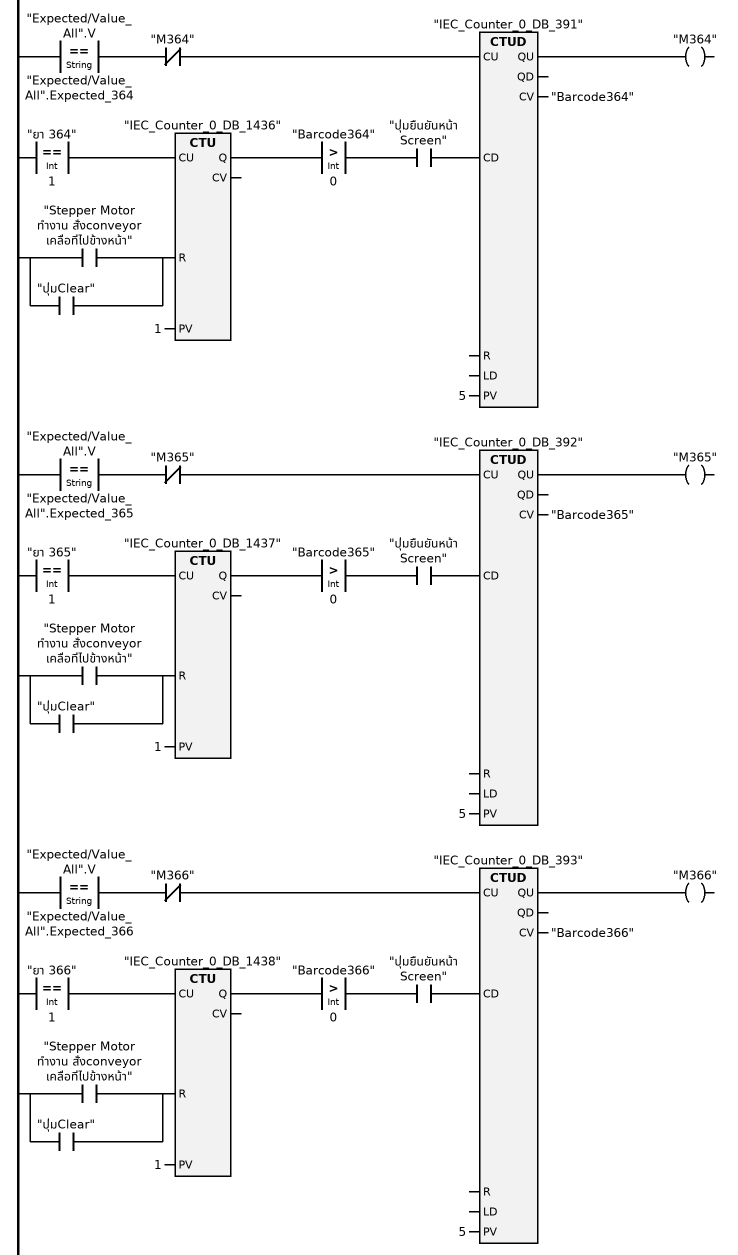
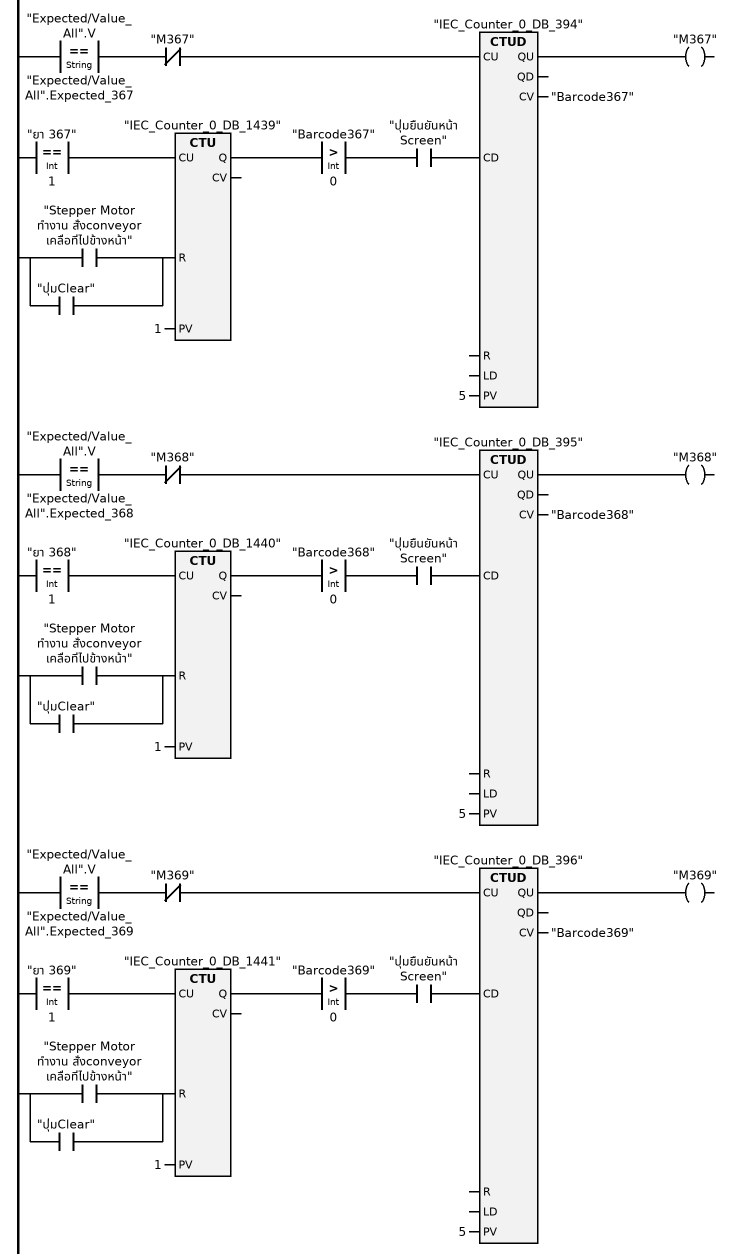
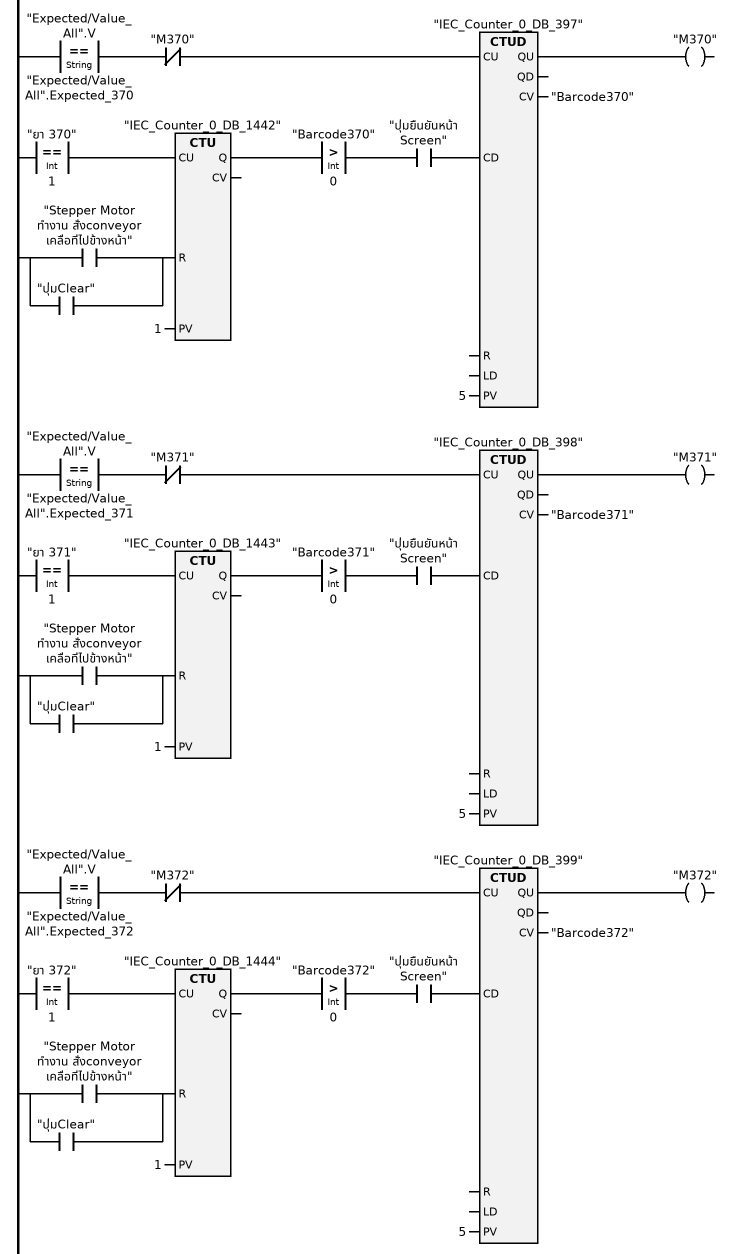
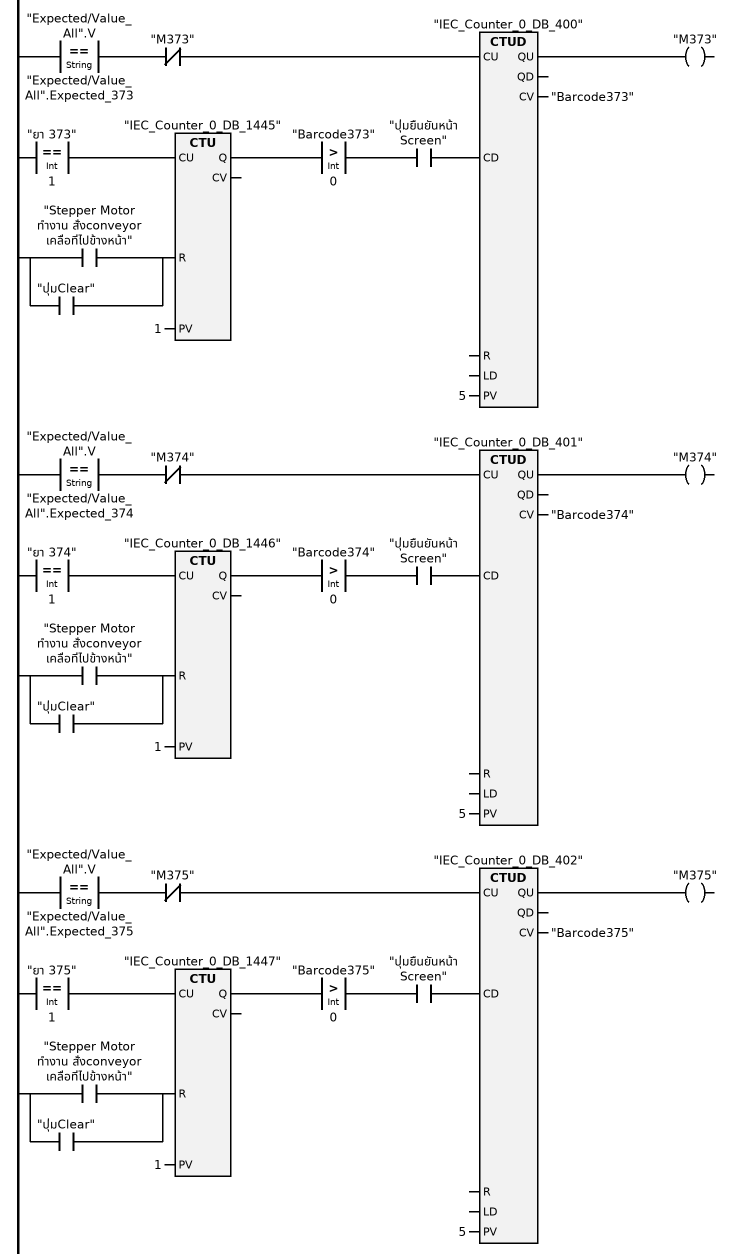
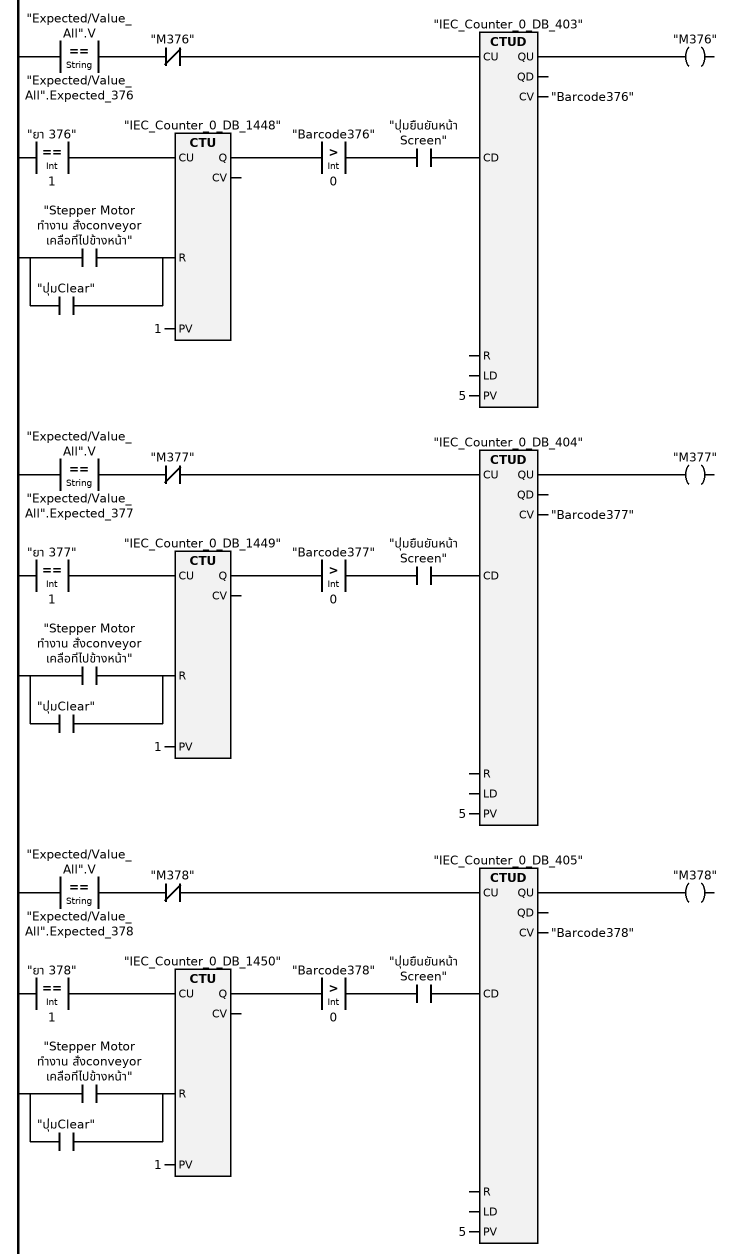
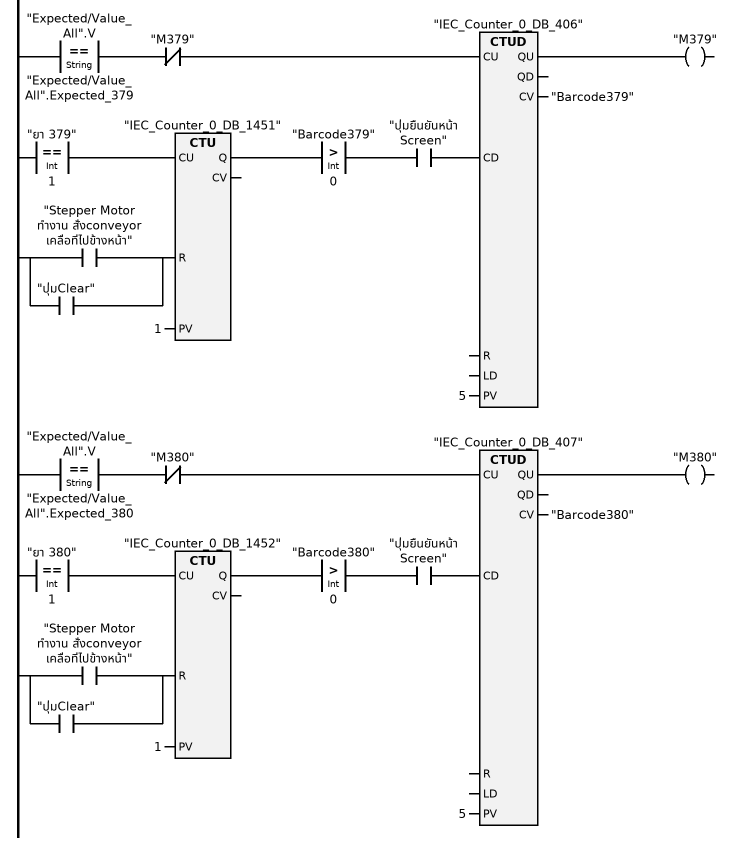
   "IEC_Counter_0_DB_1433".CTU(CU := "ยา 361" = 1,
                           R := "Stepper Motor ทำงาน สั่งconveyor เคลื่อที่ไปข้างหน้า" OR "ปุ่มClear",
                           PV := 1);
   "IEC_Counter_0_DB_388".CTUD(CU := ("Expected/Value_All".V = "Expected/Value_All".Expected_361) AND NOT "M361",
                           CD := "IEC_Counter_0_DB_1433".Q AND ("Barcode361" > 0) AND "ปุ่มยืนยันหน้า Screen",
                           PV := 5,
                           CV => "Barcode361");
   "M361" := "IEC_Counter_0_DB_388".QU;
   "IEC_Counter_0_DB_1434".CTU(CU := "ยา 362" = 1,
                           R := "Stepper Motor ทำงาน สั่งconveyor เคลื่อที่ไปข้างหน้า" OR "ปุ่มClear",
                           PV := 1);
   "IEC_Counter_0_DB_389".CTUD(CU := ("Expected/Value_All".V = "Expected/Value_All".Expected_362) AND NOT "M362",
                           CD := "IEC_Counter_0_DB_1434".Q AND ("Barcode362" > 0) AND "ปุ่มยืนยันหน้า Screen",
                           PV := 5,
                           CV => "Barcode362");
   "M362" := "IEC_Counter_0_DB_389".QU;
   "IEC_Counter_0_DB_1435".CTU(CU := "ยา 363" = 1,
                           R := "Stepper Motor ทำงาน สั่งconveyor เคลื่อที่ไปข้างหน้า" OR "ปุ่มClear",
                           PV := 1);
   "IEC_Counter_0_DB_390".CTUD(CU := ("Expected/Value_All".V = "Expected/Value_All".Expected_363) AND NOT "M363",
                           CD := "IEC_Counter_0_DB_1435".Q AND ("Barcode363" > 0) AND "ปุ่มยืนยันหน้า Screen",
                           PV := 5,
                           CV => "Barcode363");
   "M363" := "IEC_Counter_0_DB_390".QU;
   "IEC_Counter_0_DB_1436".CTU(CU := "ยา 364" = 1,
                           R := "Stepper Motor ทำงาน สั่งconveyor เคลื่อที่ไปข้างหน้า" OR "ปุ่มClear",
                           PV := 1);
   "IEC_Counter_0_DB_391".CTUD(CU := ("Expected/Value_All".V = "Expected/Value_All".Expected_364) AND NOT "M364",
                           CD := "IEC_Counter_0_DB_1436".Q AND ("Barcode364" > 0) AND "ปุ่มยืนยันหน้า Screen",
                           PV := 5,
                           CV => "Barcode364");
   "M364" := "IEC_Counter_0_DB_391".QU;
   "IEC_Counter_0_DB_1437".CTU(CU := "ยา 365" = 1,
                           R := "Stepper Motor ทำงาน สั่งconveyor เคลื่อที่ไปข้างหน้า" OR "ปุ่มClear",
                           PV := 1);
   "IEC_Counter_0_DB_392".CTUD(CU := ("Expected/Value_All".V = "Expected/Value_All".Expected_365) AND NOT "M365",
                           CD := "IEC_Counter_0_DB_1437".Q AND ("Barcode365" > 0) AND "ปุ่มยืนยันหน้า Screen",
                           PV := 5,
                           CV => "Barcode365");
   "M365" := "IEC_Counter_0_DB_392".QU;
   "IEC_Counter_0_DB_1438".CTU(CU := "ยา 366" = 1,
                           R := "Stepper Motor ทำงาน สั่งconveyor เคลื่อที่ไปข้างหน้า" OR "ปุ่มClear",
                           PV := 1);
   "IEC_Counter_0_DB_393".CTUD(CU := ("Expected/Value_All".V = "Expected/Value_All".Expected_366) AND NOT "M366",
                           CD := "IEC_Counter_0_DB_1438".Q AND ("Barcode366" > 0) AND "ปุ่มยืนยันหน้า Screen",
                           PV := 5,
                           CV => "Barcode366");
   "M366" := "IEC_Counter_0_DB_393".QU;
   "IEC_Counter_0_DB_1439".CTU(CU := "ยา 367" = 1,
                           R := "Stepper Motor ทำงาน สั่งconveyor เคลื่อที่ไปข้างหน้า" OR "ปุ่มClear",
                           PV := 1);
   "IEC_Counter_0_DB_394".CTUD(CU := ("Expected/Value_All".V = "Expected/Value_All".Expected_367) AND NOT "M367",
                           CD := "IEC_Counter_0_DB_1439".Q AND ("Barcode367" > 0) AND "ปุ่มยืนยันหน้า Screen",
                           PV := 5,
                           CV => "Barcode367");
   "M367" := "IEC_Counter_0_DB_394".QU;
   "IEC_Counter_0_DB_1440".CTU(CU := "ยา 368" = 1,
                           R := "Stepper Motor ทำงาน สั่งconveyor เคลื่อที่ไปข้างหน้า" OR "ปุ่มClear",
                           PV := 1);
   "IEC_Counter_0_DB_395".CTUD(CU := ("Expected/Value_All".V = "Expected/Value_All".Expected_368) AND NOT "M368",
                           CD := "IEC_Counter_0_DB_1440".Q AND ("Barcode368" > 0) AND "ปุ่มยืนยันหน้า Screen",
                           PV := 5,
                           CV => "Barcode368");
   "M368" := "IEC_Counter_0_DB_395".QU;
   "IEC_Counter_0_DB_1441".CTU(CU := "ยา 369" = 1,
                           R := "Stepper Motor ทำงาน สั่งconveyor เคลื่อที่ไปข้างหน้า" OR "ปุ่มClear",
                           PV := 1);
   "IEC_Counter_0_DB_396".CTUD(CU := ("Expected/Value_All".V = "Expected/Value_All".Expected_369) AND NOT "M369",
                           CD := "IEC_Counter_0_DB_1441".Q AND ("Barcode369" > 0) AND "ปุ่มยืนยันหน้า Screen",
                           PV := 5,
                           CV => "Barcode369");
   "M369" := "IEC_Counter_0_DB_396".QU;
   "IEC_Counter_0_DB_1442".CTU(CU := "ยา 370" = 1,
                           R := "Stepper Motor ทำงาน สั่งconveyor เคลื่อที่ไปข้างหน้า" OR "ปุ่มClear",
                           PV := 1);
   "IEC_Counter_0_DB_397".CTUD(CU := ("Expected/Value_All".V = "Expected/Value_All".Expected_370) AND NOT "M370",
                           CD := "IEC_Counter_0_DB_1442".Q AND ("Barcode370" > 0) AND "ปุ่มยืนยันหน้า Screen",
                           PV := 5,
                           CV => "Barcode370");
   "M370" := "IEC_Counter_0_DB_397".QU;
   "IEC_Counter_0_DB_1443".CTU(CU := "ยา 371" = 1,
                           R := "Stepper Motor ทำงาน สั่งconveyor เคลื่อที่ไปข้างหน้า" OR "ปุ่มClear",
                           PV := 1);
   "IEC_Counter_0_DB_398".CTUD(CU := ("Expected/Value_All".V = "Expected/Value_All".Expected_371) AND NOT "M371",
                           CD := "IEC_Counter_0_DB_1443".Q AND ("Barcode371" > 0) AND "ปุ่มยืนยันหน้า Screen",
                           PV := 5,
                           CV => "Barcode371");
   "M371" := "IEC_Counter_0_DB_398".QU;
   "IEC_Counter_0_DB_1444".CTU(CU := "ยา 372" = 1,
                           R := "Stepper Motor ทำงาน สั่งconveyor เคลื่อที่ไปข้างหน้า" OR "ปุ่มClear",
                           PV := 1);
   "IEC_Counter_0_DB_399".CTUD(CU := ("Expected/Value_All".V = "Expected/Value_All".Expected_372) AND NOT "M372",
                           CD := "IEC_Counter_0_DB_1444".Q AND ("Barcode372" > 0) AND "ปุ่มยืนยันหน้า Screen",
                           PV := 5,
                           CV => "Barcode372");
   "M372" := "IEC_Counter_0_DB_399".QU;
   "IEC_Counter_0_DB_1445".CTU(CU := "ยา 373" = 1,
                           R := "Stepper Motor ทำงาน สั่งconveyor เคลื่อที่ไปข้างหน้า" OR "ปุ่มClear",
                           PV := 1);
   "IEC_Counter_0_DB_400".CTUD(CU := ("Expected/Value_All".V = "Expected/Value_All".Expected_373) AND NOT "M373",
                           CD := "IEC_Counter_0_DB_1445".Q AND ("Barcode373" > 0) AND "ปุ่มยืนยันหน้า Screen",
                           PV := 5,
                           CV => "Barcode373");
   "M373" := "IEC_Counter_0_DB_400".QU;
   "IEC_Counter_0_DB_1446".CTU(CU := "ยา 374" = 1,
                           R := "Stepper Motor ทำงาน สั่งconveyor เคลื่อที่ไปข้างหน้า" OR "ปุ่มClear",
                           PV := 1);
   "IEC_Counter_0_DB_401".CTUD(CU := ("Expected/Value_All".V = "Expected/Value_All".Expected_374) AND NOT "M374",
                           CD := "IEC_Counter_0_DB_1446".Q AND ("Barcode374" > 0) AND "ปุ่มยืนยันหน้า Screen",
                           PV := 5,
                           CV => "Barcode374");
   "M374" := "IEC_Counter_0_DB_401".QU;
   "IEC_Counter_0_DB_1447".CTU(CU := "ยา 375" = 1,
                           R := "Stepper Motor ทำงาน สั่งconveyor เคลื่อที่ไปข้างหน้า" OR "ปุ่มClear",
                           PV := 1);
   "IEC_Counter_0_DB_402".CTUD(CU := ("Expected/Value_All".V = "Expected/Value_All".Expected_375) AND NOT "M375",
                           CD := "IEC_Counter_0_DB_1447".Q AND ("Barcode375" > 0) AND "ปุ่มยืนยันหน้า Screen",
                           PV := 5,
                           CV => "Barcode375");
   "M375" := "IEC_Counter_0_DB_402".QU;
   "IEC_Counter_0_DB_1448".CTU(CU := "ยา 376" = 1,
                           R := "Stepper Motor ทำงาน สั่งconveyor เคลื่อที่ไปข้างหน้า" OR "ปุ่มClear",
                           PV := 1);
   "IEC_Counter_0_DB_403".CTUD(CU := ("Expected/Value_All".V = "Expected/Value_All".Expected_376) AND NOT "M376",
                           CD := "IEC_Counter_0_DB_1448".Q AND ("Barcode376" > 0) AND "ปุ่มยืนยันหน้า Screen",
                           PV := 5,
                           CV => "Barcode376");
   "M376" := "IEC_Counter_0_DB_403".QU;
   "IEC_Counter_0_DB_1449".CTU(CU := "ยา 377" = 1,
                           R := "Stepper Motor ทำงาน สั่งconveyor เคลื่อที่ไปข้างหน้า" OR "ปุ่มClear",
                           PV := 1);
   "IEC_Counter_0_DB_404".CTUD(CU := ("Expected/Value_All".V = "Expected/Value_All".Expected_377) AND NOT "M377",
                           CD := "IEC_Counter_0_DB_1449".Q AND ("Barcode377" > 0) AND "ปุ่มยืนยันหน้า Screen",
                           PV := 5,
                           CV => "Barcode377");
   "M377" := "IEC_Counter_0_DB_404".QU;
   "IEC_Counter_0_DB_1450".CTU(CU := "ยา 378" = 1,
                           R := "Stepper Motor ทำงาน สั่งconveyor เคลื่อที่ไปข้างหน้า" OR "ปุ่มClear",
                           PV := 1);
   "IEC_Counter_0_DB_405".CTUD(CU := ("Expected/Value_All".V = "Expected/Value_All".Expected_378) AND NOT "M378",
                           CD := "IEC_Counter_0_DB_1450".Q AND ("Barcode378" > 0) AND "ปุ่มยืนยันหน้า Screen",
                           PV := 5,
                           CV => "Barcode378");
   "M378" := "IEC_Counter_0_DB_405".QU;
   "IEC_Counter_0_DB_1451".CTU(CU := "ยา 379" = 1,
                           R := "Stepper Motor ทำงาน สั่งconveyor เคลื่อที่ไปข้างหน้า" OR "ปุ่มClear",
                           PV := 1);
   "IEC_Counter_0_DB_406".CTUD(CU := ("Expected/Value_All".V = "Expected/Value_All".Expected_379) AND NOT "M379",
                           CD := "IEC_Counter_0_DB_1451".Q AND ("Barcode379" > 0) AND "ปุ่มยืนยันหน้า Screen",
                           PV := 5,
                           CV => "Barcode379");
   "M379" := "IEC_Counter_0_DB_406".QU;
   "IEC_Counter_0_DB_1452".CTU(CU := "ยา 380" = 1,
                           R := "Stepper Motor ทำงาน สั่งconveyor เคลื่อที่ไปข้างหน้า" OR "ปุ่มClear",
                           PV := 1);
   "IEC_Counter_0_DB_407".CTUD(CU := ("Expected/Value_All".V = "Expected/Value_All".Expected_380) AND NOT "M380",
                           CD := "IEC_Counter_0_DB_1452".Q AND ("Barcode380" > 0) AND "ปุ่มยืนยันหน้า Screen",
                           PV := 5,
                           CV => "Barcode380");
   "M380" := "IEC_Counter_0_DB_407".QU;
END_REGION

REGION Network 20
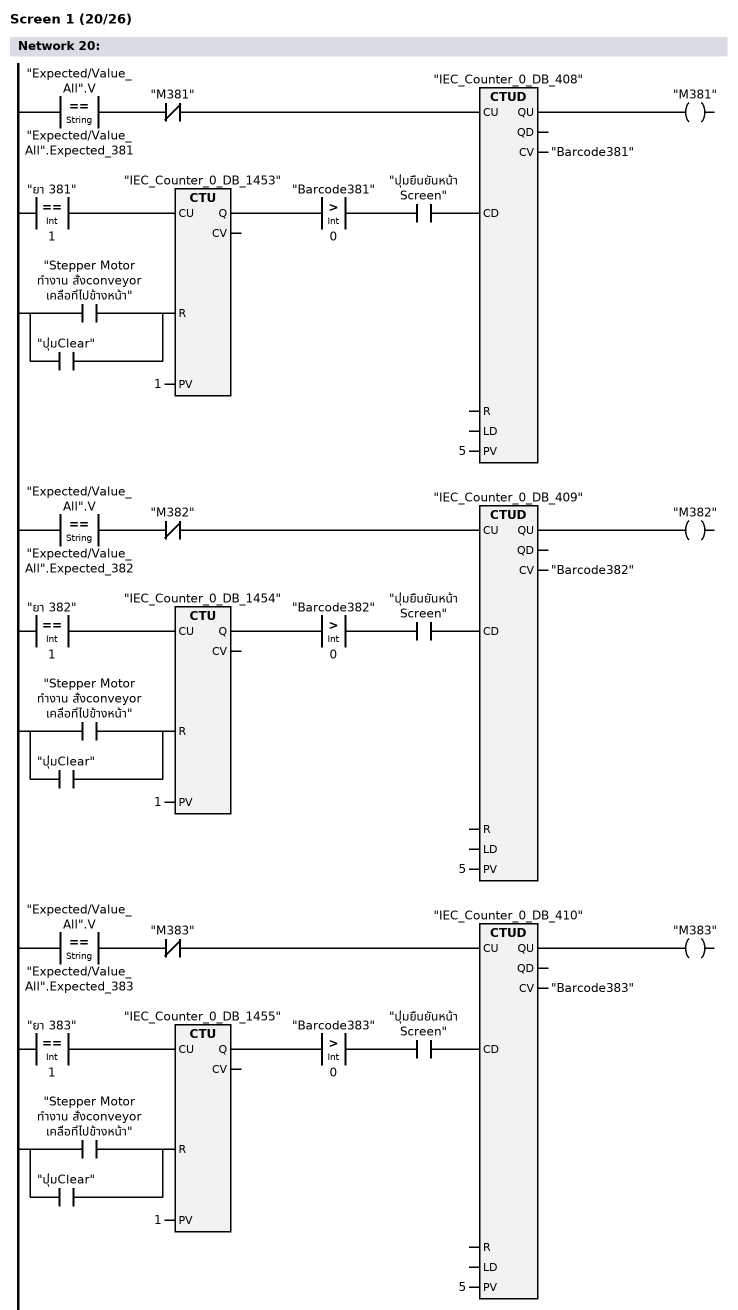
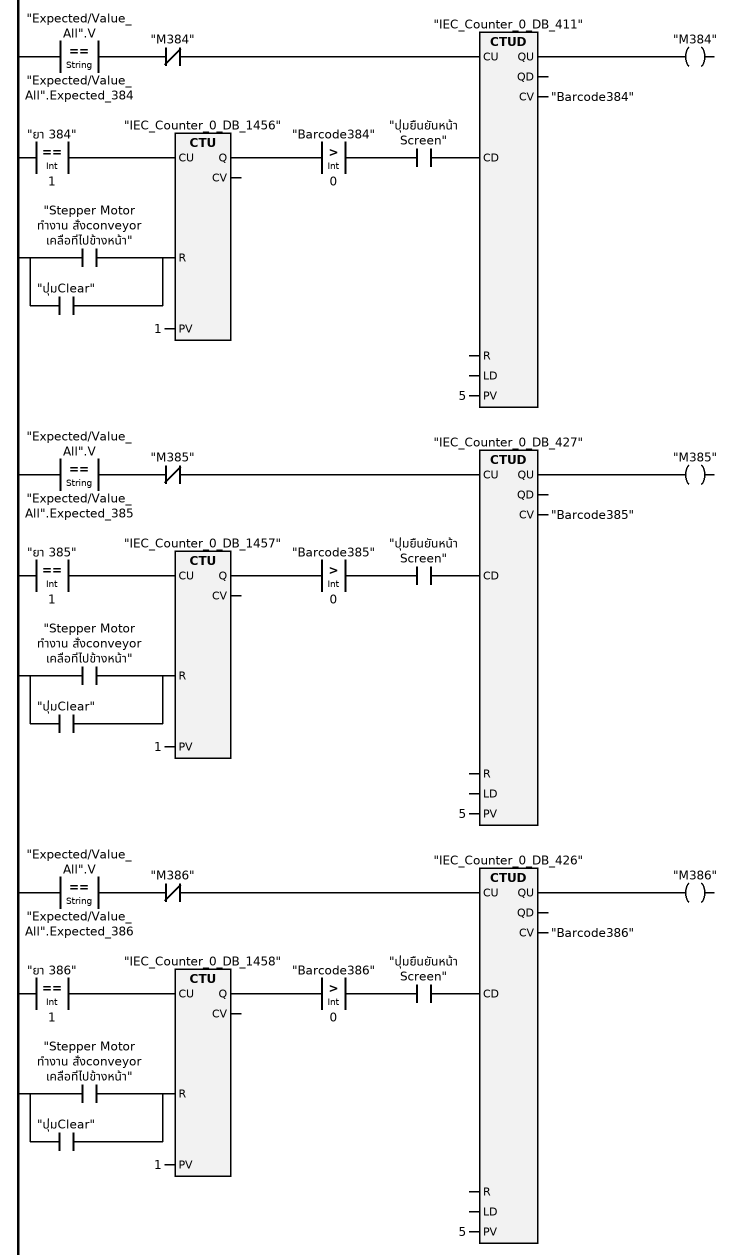
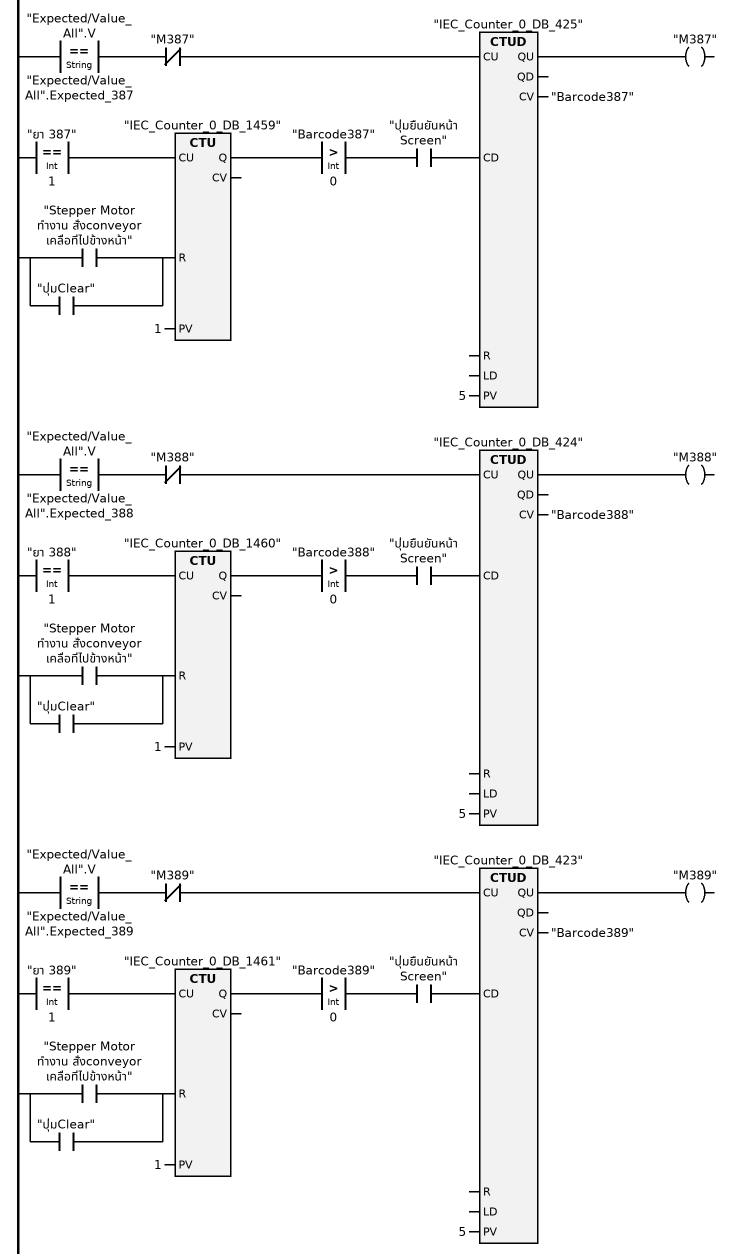
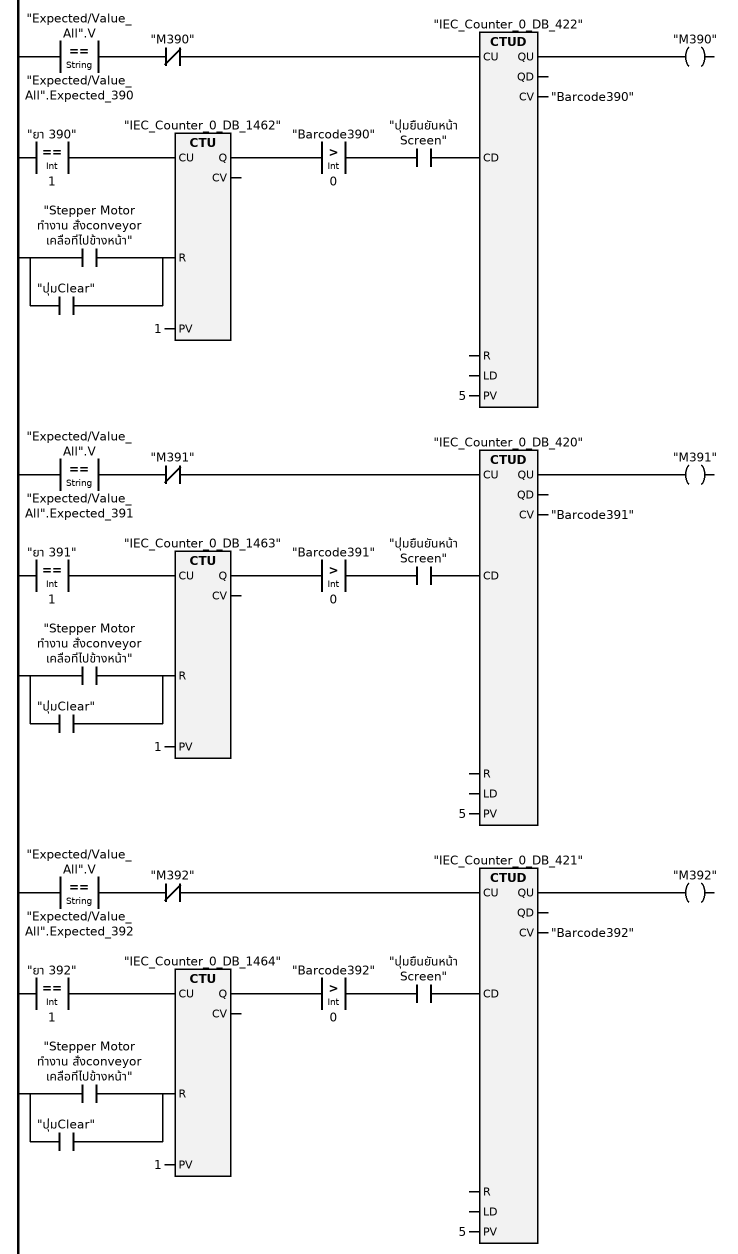
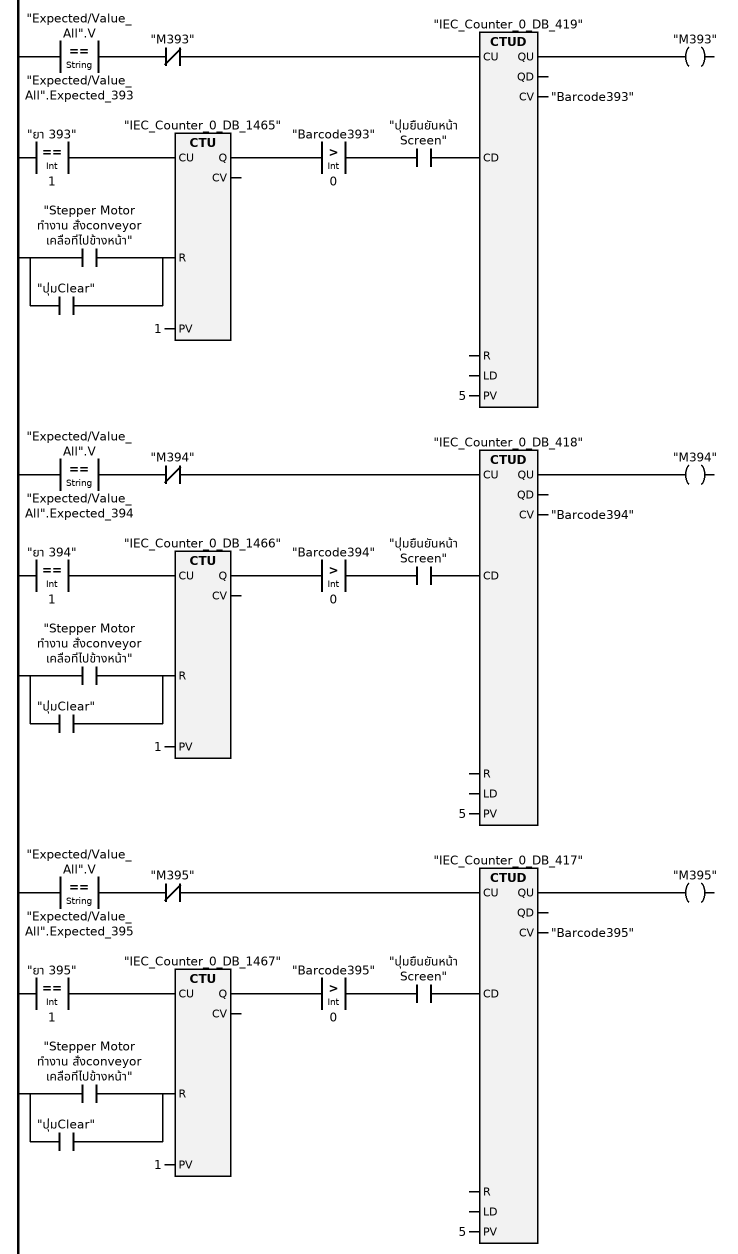
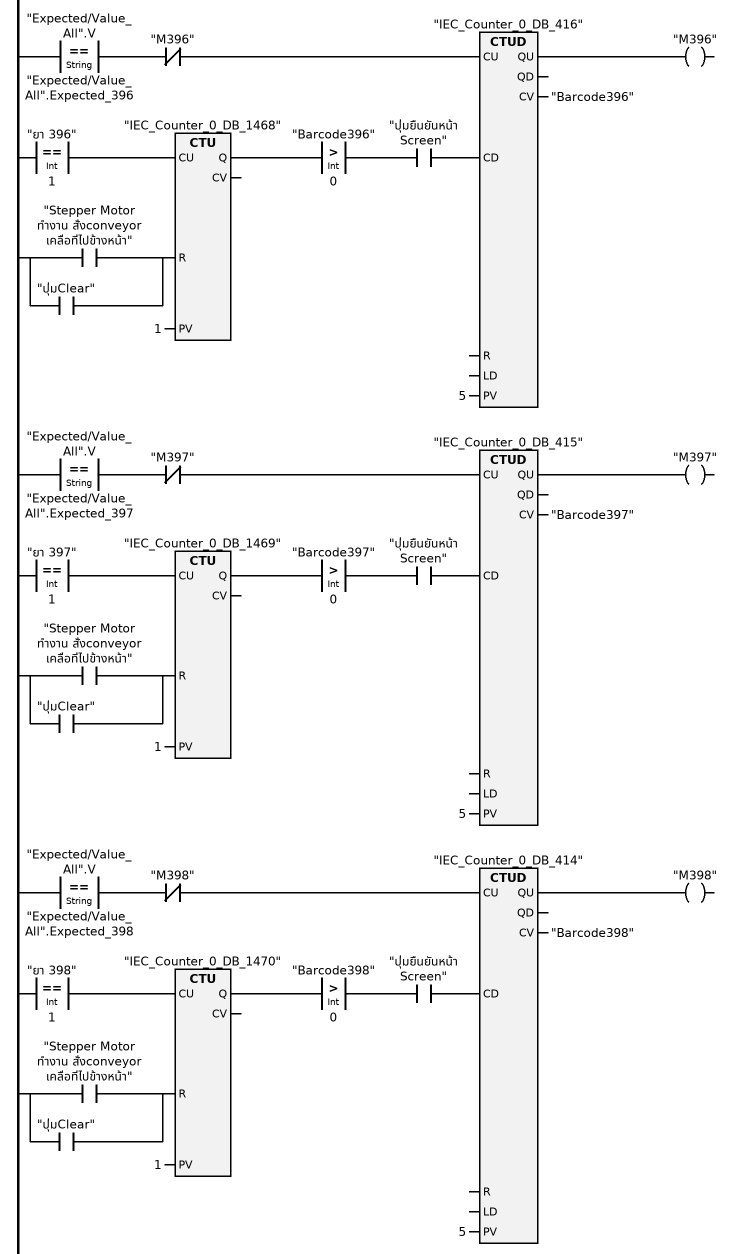
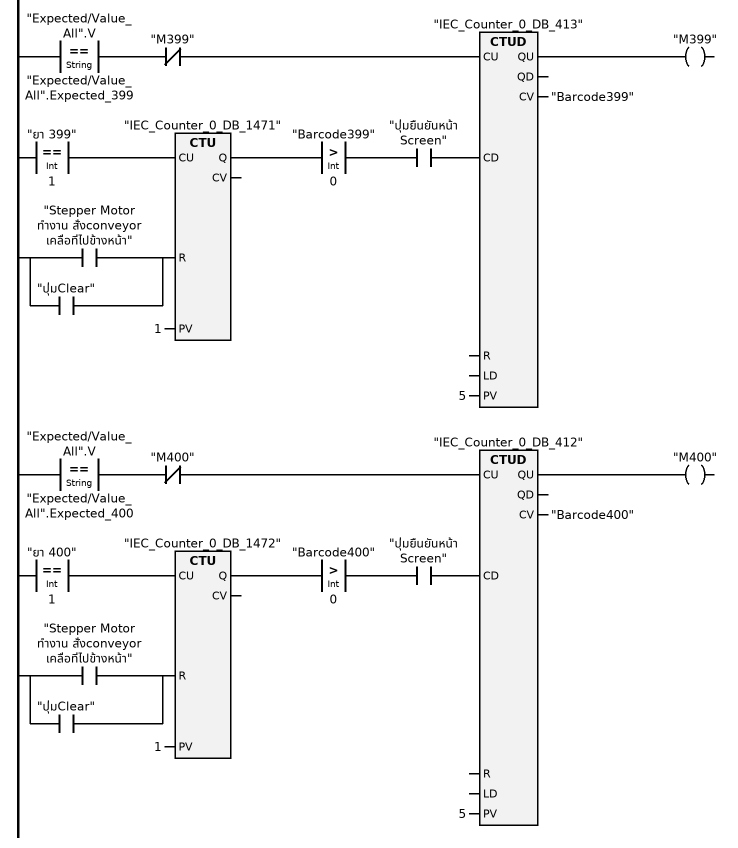
   "IEC_Counter_0_DB_1453".CTU(CU := "ยา 381" = 1,
                           R := "Stepper Motor ทำงาน สั่งconveyor เคลื่อที่ไปข้างหน้า" OR "ปุ่มClear",
                           PV := 1);
   "IEC_Counter_0_DB_408".CTUD(CU := ("Expected/Value_All".V = "Expected/Value_All".Expected_381) AND NOT "M381",
                           CD := "IEC_Counter_0_DB_1453".Q AND ("Barcode381" > 0) AND "ปุ่มยืนยันหน้า Screen",
                           PV := 5,
                           CV => "Barcode381");
   "M381" := "IEC_Counter_0_DB_408".QU;
   "IEC_Counter_0_DB_1454".CTU(CU := "ยา 382" = 1,
                           R := "Stepper Motor ทำงาน สั่งconveyor เคลื่อที่ไปข้างหน้า" OR "ปุ่มClear",
                           PV := 1);
   "IEC_Counter_0_DB_409".CTUD(CU := ("Expected/Value_All".V = "Expected/Value_All".Expected_382) AND NOT "M382",
                           CD := "IEC_Counter_0_DB_1454".Q AND ("Barcode382" > 0) AND "ปุ่มยืนยันหน้า Screen",
                           PV := 5,
                           CV => "Barcode382");
   "M382" := "IEC_Counter_0_DB_409".QU;
   "IEC_Counter_0_DB_1455".CTU(CU := "ยา 383" = 1,
                           R := "Stepper Motor ทำงาน สั่งconveyor เคลื่อที่ไปข้างหน้า" OR "ปุ่มClear",
                           PV := 1);
   "IEC_Counter_0_DB_410".CTUD(CU := ("Expected/Value_All".V = "Expected/Value_All".Expected_383) AND NOT "M383",
                           CD := "IEC_Counter_0_DB_1455".Q AND ("Barcode383" > 0) AND "ปุ่มยืนยันหน้า Screen",
                           PV := 5,
                           CV => "Barcode383");
   "M383" := "IEC_Counter_0_DB_410".QU;
   "IEC_Counter_0_DB_1456".CTU(CU := "ยา 384" = 1,
                           R := "Stepper Motor ทำงาน สั่งconveyor เคลื่อที่ไปข้างหน้า" OR "ปุ่มClear",
                           PV := 1);
   "IEC_Counter_0_DB_411".CTUD(CU := ("Expected/Value_All".V = "Expected/Value_All".Expected_384) AND NOT "M384",
                           CD := "IEC_Counter_0_DB_1456".Q AND ("Barcode384" > 0) AND "ปุ่มยืนยันหน้า Screen",
                           PV := 5,
                           CV => "Barcode384");
   "M384" := "IEC_Counter_0_DB_411".QU;
   "IEC_Counter_0_DB_1457".CTU(CU := "ยา 385" = 1,
                           R := "Stepper Motor ทำงาน สั่งconveyor เคลื่อที่ไปข้างหน้า" OR "ปุ่มClear",
                           PV := 1);
   "IEC_Counter_0_DB_427".CTUD(CU := ("Expected/Value_All".V = "Expected/Value_All".Expected_385) AND NOT "M385",
                           CD := "IEC_Counter_0_DB_1457".Q AND ("Barcode385" > 0) AND "ปุ่มยืนยันหน้า Screen",
                           PV := 5,
                           CV => "Barcode385");
   "M385" := "IEC_Counter_0_DB_427".QU;
   "IEC_Counter_0_DB_1458".CTU(CU := "ยา 386" = 1,
                           R := "Stepper Motor ทำงาน สั่งconveyor เคลื่อที่ไปข้างหน้า" OR "ปุ่มClear",
                           PV := 1);
   "IEC_Counter_0_DB_426".CTUD(CU := ("Expected/Value_All".V = "Expected/Value_All".Expected_386) AND NOT "M386",
                           CD := "IEC_Counter_0_DB_1458".Q AND ("Barcode386" > 0) AND "ปุ่มยืนยันหน้า Screen",
                           PV := 5,
                           CV => "Barcode386");
   "M386" := "IEC_Counter_0_DB_426".QU;
   "IEC_Counter_0_DB_1459".CTU(CU := "ยา 387" = 1,
                           R := "Stepper Motor ทำงาน สั่งconveyor เคลื่อที่ไปข้างหน้า" OR "ปุ่มClear",
                           PV := 1);
   "IEC_Counter_0_DB_425".CTUD(CU := ("Expected/Value_All".V = "Expected/Value_All".Expected_387) AND NOT "M387",
                           CD := "IEC_Counter_0_DB_1459".Q AND ("Barcode387" > 0) AND "ปุ่มยืนยันหน้า Screen",
                           PV := 5,
                           CV => "Barcode387");
   "M387" := "IEC_Counter_0_DB_425".QU;
   "IEC_Counter_0_DB_1460".CTU(CU := "ยา 388" = 1,
                           R := "Stepper Motor ทำงาน สั่งconveyor เคลื่อที่ไปข้างหน้า" OR "ปุ่มClear",
                           PV := 1);
   "IEC_Counter_0_DB_424".CTUD(CU := ("Expected/Value_All".V = "Expected/Value_All".Expected_388) AND NOT "M388",
                           CD := "IEC_Counter_0_DB_1460".Q AND ("Barcode388" > 0) AND "ปุ่มยืนยันหน้า Screen",
                           PV := 5,
                           CV => "Barcode388");
   "M388" := "IEC_Counter_0_DB_424".QU;
   "IEC_Counter_0_DB_1461".CTU(CU := "ยา 389" = 1,
                           R := "Stepper Motor ทำงาน สั่งconveyor เคลื่อที่ไปข้างหน้า" OR "ปุ่มClear",
                           PV := 1);
   "IEC_Counter_0_DB_423".CTUD(CU := ("Expected/Value_All".V = "Expected/Value_All".Expected_389) AND NOT "M389",
                           CD := "IEC_Counter_0_DB_1461".Q AND ("Barcode389" > 0) AND "ปุ่มยืนยันหน้า Screen",
                           PV := 5,
                           CV => "Barcode389");
   "M389" := "IEC_Counter_0_DB_423".QU;
   "IEC_Counter_0_DB_1462".CTU(CU := "ยา 390" = 1,
                           R := "Stepper Motor ทำงาน สั่งconveyor เคลื่อที่ไปข้างหน้า" OR "ปุ่มClear",
                           PV := 1);
   "IEC_Counter_0_DB_422".CTUD(CU := ("Expected/Value_All".V = "Expected/Value_All".Expected_390) AND NOT "M390",
                           CD := "IEC_Counter_0_DB_1462".Q AND ("Barcode390" > 0) AND "ปุ่มยืนยันหน้า Screen",
                           PV := 5,
                           CV => "Barcode390");
   "M390" := "IEC_Counter_0_DB_422".QU;
   "IEC_Counter_0_DB_1463".CTU(CU := "ยา 391" = 1,
                           R := "Stepper Motor ทำงาน สั่งconveyor เคลื่อที่ไปข้างหน้า" OR "ปุ่มClear",
                           PV := 1);
   "IEC_Counter_0_DB_420".CTUD(CU := ("Expected/Value_All".V = "Expected/Value_All".Expected_391) AND NOT "M391",
                           CD := "IEC_Counter_0_DB_1463".Q AND ("Barcode391" > 0) AND "ปุ่มยืนยันหน้า Screen",
                           PV := 5,
                           CV => "Barcode391");
   "M391" := "IEC_Counter_0_DB_420".QU;
   "IEC_Counter_0_DB_1464".CTU(CU := "ยา 392" = 1,
                           R := "Stepper Motor ทำงาน สั่งconveyor เคลื่อที่ไปข้างหน้า" OR "ปุ่มClear",
                           PV := 1);
   "IEC_Counter_0_DB_421".CTUD(CU := ("Expected/Value_All".V = "Expected/Value_All".Expected_392) AND NOT "M392",
                           CD := "IEC_Counter_0_DB_1464".Q AND ("Barcode392" > 0) AND "ปุ่มยืนยันหน้า Screen",
                           PV := 5,
                           CV => "Barcode392");
   "M392" := "IEC_Counter_0_DB_421".QU;
   "IEC_Counter_0_DB_1465".CTU(CU := "ยา 393" = 1,
                           R := "Stepper Motor ทำงาน สั่งconveyor เคลื่อที่ไปข้างหน้า" OR "ปุ่มClear",
                           PV := 1);
   "IEC_Counter_0_DB_419".CTUD(CU := ("Expected/Value_All".V = "Expected/Value_All".Expected_393) AND NOT "M393",
                           CD := "IEC_Counter_0_DB_1465".Q AND ("Barcode393" > 0) AND "ปุ่มยืนยันหน้า Screen",
                           PV := 5,
                           CV => "Barcode393");
   "M393" := "IEC_Counter_0_DB_419".QU;
   "IEC_Counter_0_DB_1466".CTU(CU := "ยา 394" = 1,
                           R := "Stepper Motor ทำงาน สั่งconveyor เคลื่อที่ไปข้างหน้า" OR "ปุ่มClear",
                           PV := 1);
   "IEC_Counter_0_DB_418".CTUD(CU := ("Expected/Value_All".V = "Expected/Value_All".Expected_394) AND NOT "M394",
                           CD := "IEC_Counter_0_DB_1466".Q AND ("Barcode394" > 0) AND "ปุ่มยืนยันหน้า Screen",
                           PV := 5,
                           CV => "Barcode394");
   "M394" := "IEC_Counter_0_DB_418".QU;
   "IEC_Counter_0_DB_1467".CTU(CU := "ยา 395" = 1,
                           R := "Stepper Motor ทำงาน สั่งconveyor เคลื่อที่ไปข้างหน้า" OR "ปุ่มClear",
                           PV := 1);
   "IEC_Counter_0_DB_417".CTUD(CU := ("Expected/Value_All".V = "Expected/Value_All".Expected_395) AND NOT "M395",
                           CD := "IEC_Counter_0_DB_1467".Q AND ("Barcode395" > 0) AND "ปุ่มยืนยันหน้า Screen",
                           PV := 5,
                           CV => "Barcode395");
   "M395" := "IEC_Counter_0_DB_417".QU;
   "IEC_Counter_0_DB_1468".CTU(CU := "ยา 396" = 1,
                           R := "Stepper Motor ทำงาน สั่งconveyor เคลื่อที่ไปข้างหน้า" OR "ปุ่มClear",
                           PV := 1);
   "IEC_Counter_0_DB_416".CTUD(CU := ("Expected/Value_All".V = "Expected/Value_All".Expected_396) AND NOT "M396",
                           CD := "IEC_Counter_0_DB_1468".Q AND ("Barcode396" > 0) AND "ปุ่มยืนยันหน้า Screen",
                           PV := 5,
                           CV => "Barcode396");
   "M396" := "IEC_Counter_0_DB_416".QU;
   "IEC_Counter_0_DB_1469".CTU(CU := "ยา 397" = 1,
                           R := "Stepper Motor ทำงาน สั่งconveyor เคลื่อที่ไปข้างหน้า" OR "ปุ่มClear",
                           PV := 1);
   "IEC_Counter_0_DB_415".CTUD(CU := ("Expected/Value_All".V = "Expected/Value_All".Expected_397) AND NOT "M397",
                           CD := "IEC_Counter_0_DB_1469".Q AND ("Barcode397" > 0) AND "ปุ่มยืนยันหน้า Screen",
                           PV := 5,
                           CV => "Barcode397");
   "M397" := "IEC_Counter_0_DB_415".QU;
   "IEC_Counter_0_DB_1470".CTU(CU := "ยา 398" = 1,
                           R := "Stepper Motor ทำงาน สั่งconveyor เคลื่อที่ไปข้างหน้า" OR "ปุ่มClear",
                           PV := 1);
   "IEC_Counter_0_DB_414".CTUD(CU := ("Expected/Value_All".V = "Expected/Value_All".Expected_398) AND NOT "M398",
                           CD := "IEC_Counter_0_DB_1470".Q AND ("Barcode398" > 0) AND "ปุ่มยืนยันหน้า Screen",
                           PV := 5,
                           CV => "Barcode398");
   "M398" := "IEC_Counter_0_DB_414".QU;
   "IEC_Counter_0_DB_1471".CTU(CU := "ยา 399" = 1,
                           R := "Stepper Motor ทำงาน สั่งconveyor เคลื่อที่ไปข้างหน้า" OR "ปุ่มClear",
                           PV := 1);
   "IEC_Counter_0_DB_413".CTUD(CU := ("Expected/Value_All".V = "Expected/Value_All".Expected_399) AND NOT "M399",
                           CD := "IEC_Counter_0_DB_1471".Q AND ("Barcode399" > 0) AND "ปุ่มยืนยันหน้า Screen",
                           PV := 5,
                           CV => "Barcode399");
   "M399" := "IEC_Counter_0_DB_413".QU;
   "IEC_Counter_0_DB_1472".CTU(CU := "ยา 400" = 1,
                           R := "Stepper Motor ทำงาน สั่งconveyor เคลื่อที่ไปข้างหน้า" OR "ปุ่มClear",
                           PV := 1);
   "IEC_Counter_0_DB_412".CTUD(CU := ("Expected/Value_All".V = "Expected/Value_All".Expected_400) AND NOT "M400",
                           CD := "IEC_Counter_0_DB_1472".Q AND ("Barcode400" > 0) AND "ปุ่มยืนยันหน้า Screen",
                           PV := 5,
                           CV => "Barcode400");
   "M400" := "IEC_Counter_0_DB_412".QU;
END_REGION

REGION Network 21
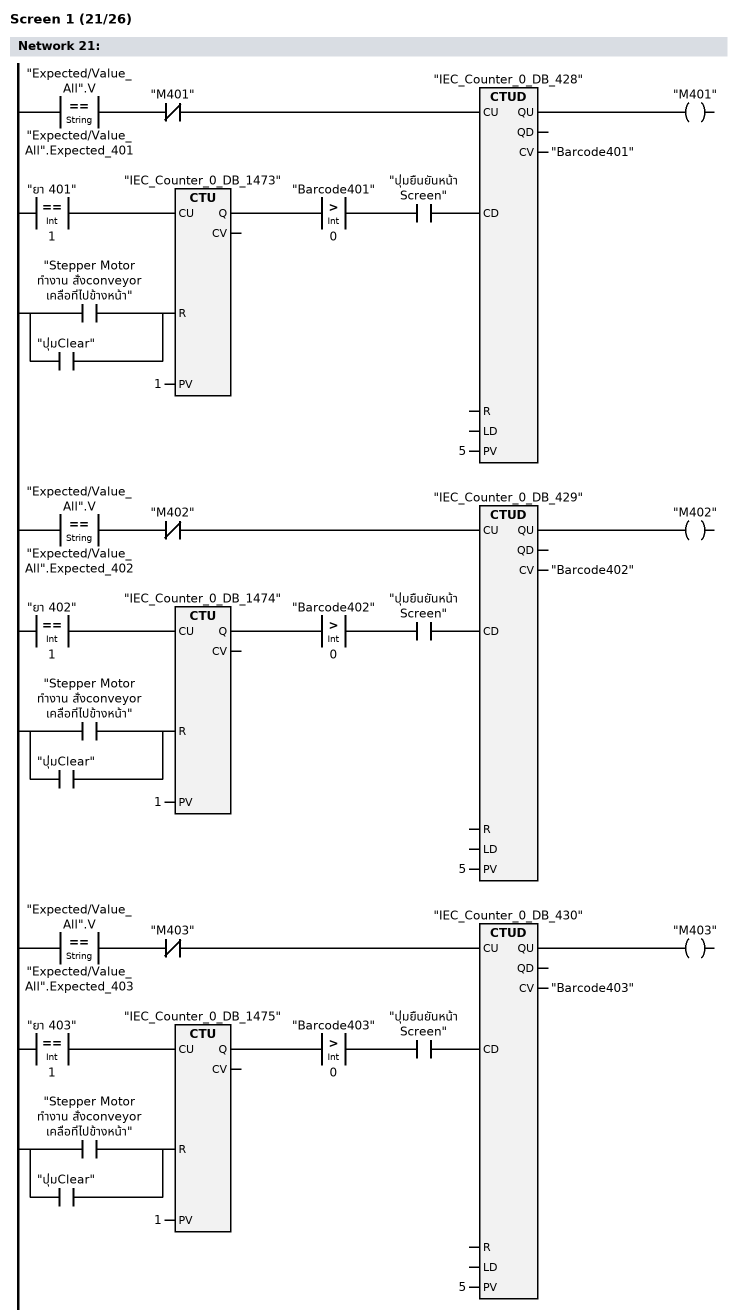
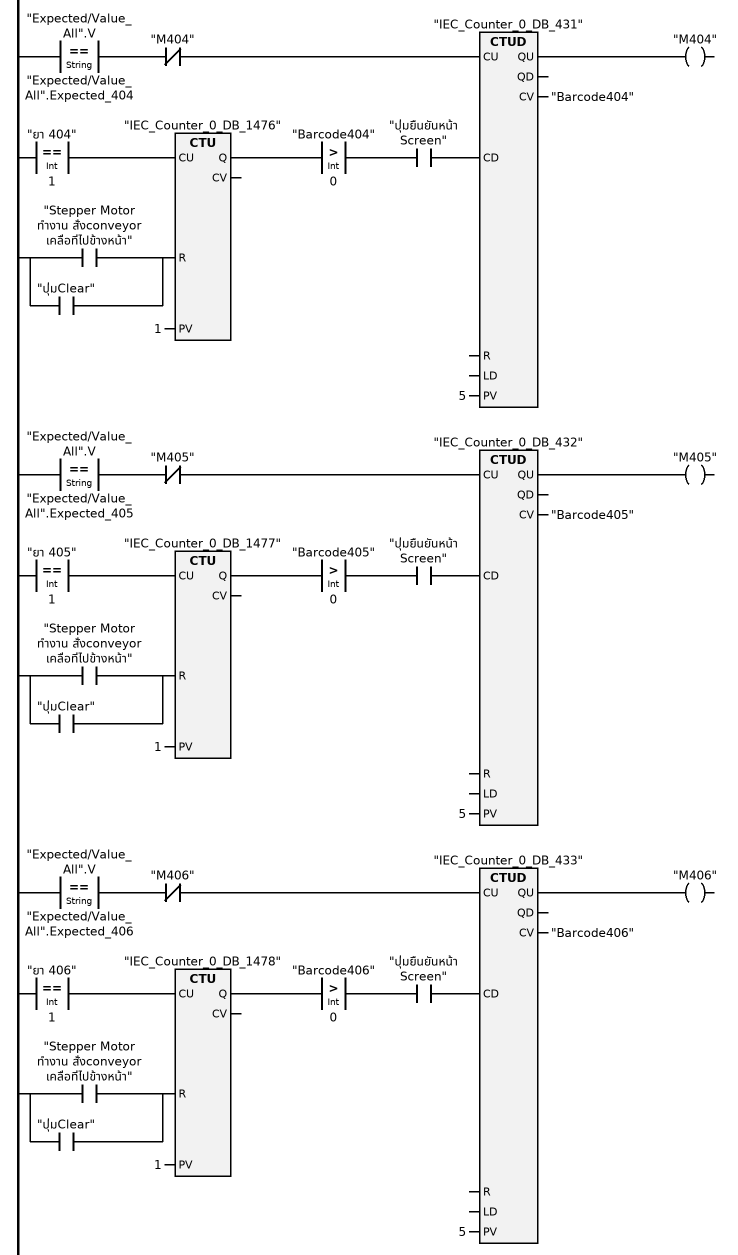
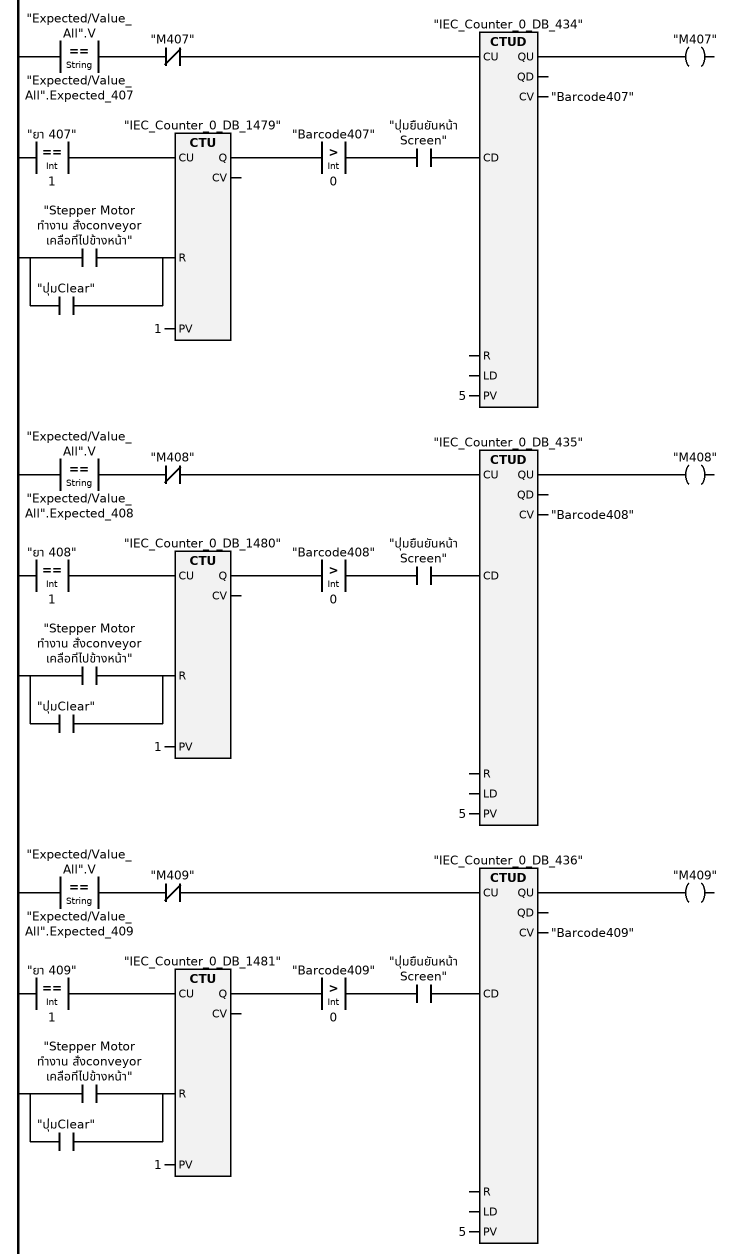
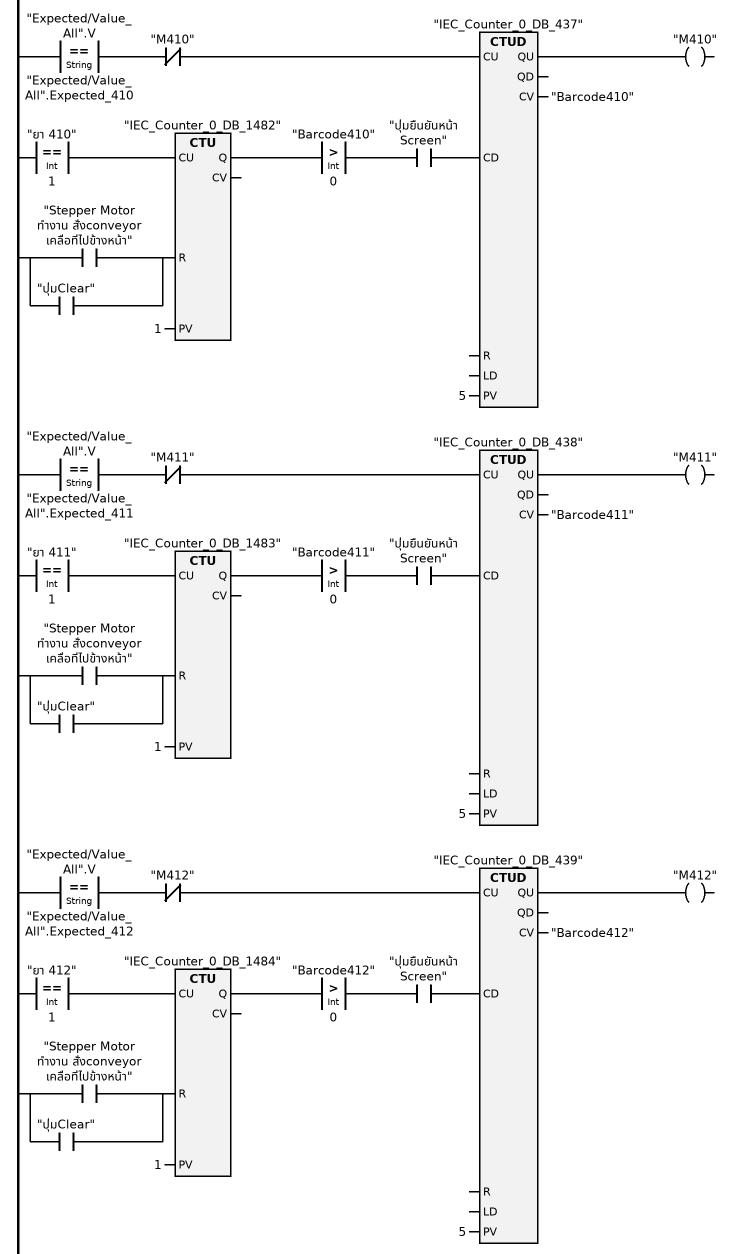
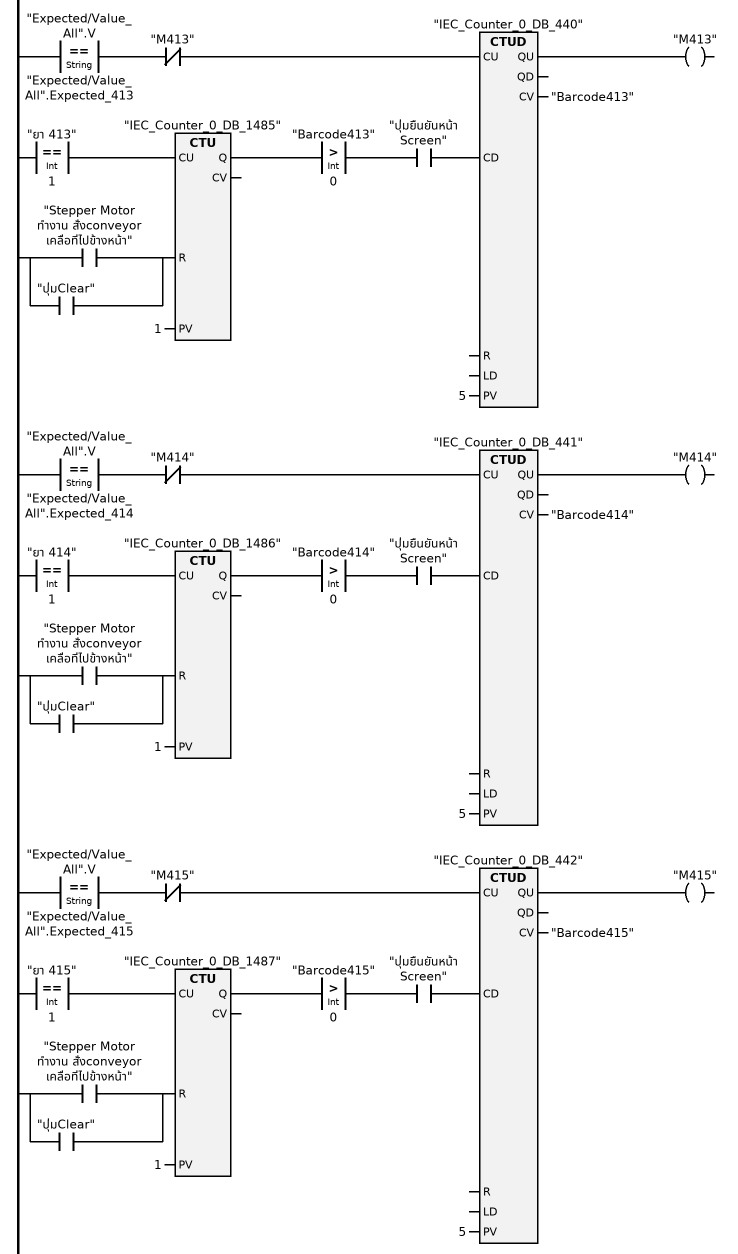
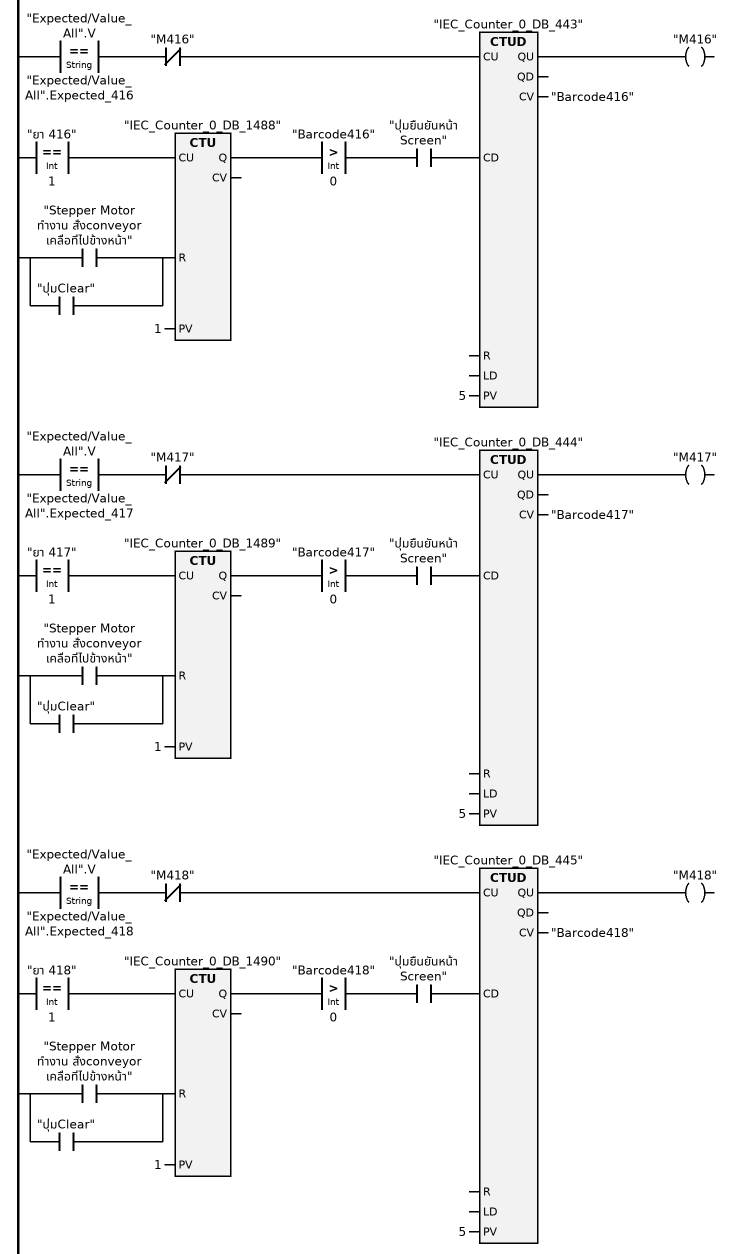
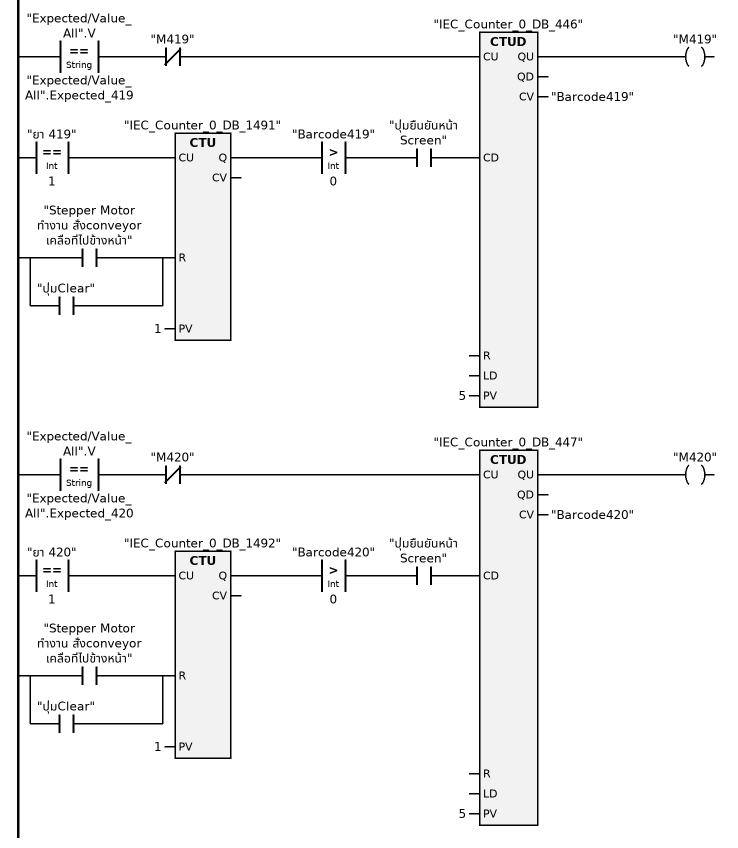
   "IEC_Counter_0_DB_1473".CTU(CU := "ยา 401" = 1,
                           R := "Stepper Motor ทำงาน สั่งconveyor เคลื่อที่ไปข้างหน้า" OR "ปุ่มClear",
                           PV := 1);
   "IEC_Counter_0_DB_428".CTUD(CU := ("Expected/Value_All".V = "Expected/Value_All".Expected_401) AND NOT "M401",
                           CD := "IEC_Counter_0_DB_1473".Q AND ("Barcode401" > 0) AND "ปุ่มยืนยันหน้า Screen",
                           PV := 5,
                           CV => "Barcode401");
   "M401" := "IEC_Counter_0_DB_428".QU;
   "IEC_Counter_0_DB_1474".CTU(CU := "ยา 402" = 1,
                           R := "Stepper Motor ทำงาน สั่งconveyor เคลื่อที่ไปข้างหน้า" OR "ปุ่มClear",
                           PV := 1);
   "IEC_Counter_0_DB_429".CTUD(CU := ("Expected/Value_All".V = "Expected/Value_All".Expected_402) AND NOT "M402",
                           CD := "IEC_Counter_0_DB_1474".Q AND ("Barcode402" > 0) AND "ปุ่มยืนยันหน้า Screen",
                           PV := 5,
                           CV => "Barcode402");
   "M402" := "IEC_Counter_0_DB_429".QU;
   "IEC_Counter_0_DB_1475".CTU(CU := "ยา 403" = 1,
                           R := "Stepper Motor ทำงาน สั่งconveyor เคลื่อที่ไปข้างหน้า" OR "ปุ่มClear",
                           PV := 1);
   "IEC_Counter_0_DB_430".CTUD(CU := ("Expected/Value_All".V = "Expected/Value_All".Expected_403) AND NOT "M403",
                           CD := "IEC_Counter_0_DB_1475".Q AND ("Barcode403" > 0) AND "ปุ่มยืนยันหน้า Screen",
                           PV := 5,
                           CV => "Barcode403");
   "M403" := "IEC_Counter_0_DB_430".QU;
   "IEC_Counter_0_DB_1476".CTU(CU := "ยา 404" = 1,
                           R := "Stepper Motor ทำงาน สั่งconveyor เคลื่อที่ไปข้างหน้า" OR "ปุ่มClear",
                           PV := 1);
   "IEC_Counter_0_DB_431".CTUD(CU := ("Expected/Value_All".V = "Expected/Value_All".Expected_404) AND NOT "M404",
                           CD := "IEC_Counter_0_DB_1476".Q AND ("Barcode404" > 0) AND "ปุ่มยืนยันหน้า Screen",
                           PV := 5,
                           CV => "Barcode404");
   "M404" := "IEC_Counter_0_DB_431".QU;
   "IEC_Counter_0_DB_1477".CTU(CU := "ยา 405" = 1,
                           R := "Stepper Motor ทำงาน สั่งconveyor เคลื่อที่ไปข้างหน้า" OR "ปุ่มClear",
                           PV := 1);
   "IEC_Counter_0_DB_432".CTUD(CU := ("Expected/Value_All".V = "Expected/Value_All".Expected_405) AND NOT "M405",
                           CD := "IEC_Counter_0_DB_1477".Q AND ("Barcode405" > 0) AND "ปุ่มยืนยันหน้า Screen",
                           PV := 5,
                           CV => "Barcode405");
   "M405" := "IEC_Counter_0_DB_432".QU;
   "IEC_Counter_0_DB_1478".CTU(CU := "ยา 406" = 1,
                           R := "Stepper Motor ทำงาน สั่งconveyor เคลื่อที่ไปข้างหน้า" OR "ปุ่มClear",
                           PV := 1);
   "IEC_Counter_0_DB_433".CTUD(CU := ("Expected/Value_All".V = "Expected/Value_All".Expected_406) AND NOT "M406",
                           CD := "IEC_Counter_0_DB_1478".Q AND ("Barcode406" > 0) AND "ปุ่มยืนยันหน้า Screen",
                           PV := 5,
                           CV => "Barcode406");
   "M406" := "IEC_Counter_0_DB_433".QU;
   "IEC_Counter_0_DB_1479".CTU(CU := "ยา 407" = 1,
                           R := "Stepper Motor ทำงาน สั่งconveyor เคลื่อที่ไปข้างหน้า" OR "ปุ่มClear",
                           PV := 1);
   "IEC_Counter_0_DB_434".CTUD(CU := ("Expected/Value_All".V = "Expected/Value_All".Expected_407) AND NOT "M407",
                           CD := "IEC_Counter_0_DB_1479".Q AND ("Barcode407" > 0) AND "ปุ่มยืนยันหน้า Screen",
                           PV := 5,
                           CV => "Barcode407");
   "M407" := "IEC_Counter_0_DB_434".QU;
   "IEC_Counter_0_DB_1480".CTU(CU := "ยา 408" = 1,
                           R := "Stepper Motor ทำงาน สั่งconveyor เคลื่อที่ไปข้างหน้า" OR "ปุ่มClear",
                           PV := 1);
   "IEC_Counter_0_DB_435".CTUD(CU := ("Expected/Value_All".V = "Expected/Value_All".Expected_408) AND NOT "M408",
                           CD := "IEC_Counter_0_DB_1480".Q AND ("Barcode408" > 0) AND "ปุ่มยืนยันหน้า Screen",
                           PV := 5,
                           CV => "Barcode408");
   "M408" := "IEC_Counter_0_DB_435".QU;
   "IEC_Counter_0_DB_1481".CTU(CU := "ยา 409" = 1,
                           R := "Stepper Motor ทำงาน สั่งconveyor เคลื่อที่ไปข้างหน้า" OR "ปุ่มClear",
                           PV := 1);
   "IEC_Counter_0_DB_436".CTUD(CU := ("Expected/Value_All".V = "Expected/Value_All".Expected_409) AND NOT "M409",
                           CD := "IEC_Counter_0_DB_1481".Q AND ("Barcode409" > 0) AND "ปุ่มยืนยันหน้า Screen",
                           PV := 5,
                           CV => "Barcode409");
   "M409" := "IEC_Counter_0_DB_436".QU;
   "IEC_Counter_0_DB_1482".CTU(CU := "ยา 410" = 1,
                           R := "Stepper Motor ทำงาน สั่งconveyor เคลื่อที่ไปข้างหน้า" OR "ปุ่มClear",
                           PV := 1);
   "IEC_Counter_0_DB_437".CTUD(CU := ("Expected/Value_All".V = "Expected/Value_All".Expected_410) AND NOT "M410",
                           CD := "IEC_Counter_0_DB_1482".Q AND ("Barcode410" > 0) AND "ปุ่มยืนยันหน้า Screen",
                           PV := 5,
                           CV => "Barcode410");
   "M410" := "IEC_Counter_0_DB_437".QU;
   "IEC_Counter_0_DB_1483".CTU(CU := "ยา 411" = 1,
                           R := "Stepper Motor ทำงาน สั่งconveyor เคลื่อที่ไปข้างหน้า" OR "ปุ่มClear",
                           PV := 1);
   "IEC_Counter_0_DB_438".CTUD(CU := ("Expected/Value_All".V = "Expected/Value_All".Expected_411) AND NOT "M411",
                           CD := "IEC_Counter_0_DB_1483".Q AND ("Barcode411" > 0) AND "ปุ่มยืนยันหน้า Screen",
                           PV := 5,
                           CV => "Barcode411");
   "M411" := "IEC_Counter_0_DB_438".QU;
   "IEC_Counter_0_DB_1484".CTU(CU := "ยา 412" = 1,
                           R := "Stepper Motor ทำงาน สั่งconveyor เคลื่อที่ไปข้างหน้า" OR "ปุ่มClear",
                           PV := 1);
   "IEC_Counter_0_DB_439".CTUD(CU := ("Expected/Value_All".V = "Expected/Value_All".Expected_412) AND NOT "M412",
                           CD := "IEC_Counter_0_DB_1484".Q AND ("Barcode412" > 0) AND "ปุ่มยืนยันหน้า Screen",
                           PV := 5,
                           CV => "Barcode412");
   "M412" := "IEC_Counter_0_DB_439".QU;
   "IEC_Counter_0_DB_1485".CTU(CU := "ยา 413" = 1,
                           R := "Stepper Motor ทำงาน สั่งconveyor เคลื่อที่ไปข้างหน้า" OR "ปุ่มClear",
                           PV := 1);
   "IEC_Counter_0_DB_440".CTUD(CU := ("Expected/Value_All".V = "Expected/Value_All".Expected_413) AND NOT "M413",
                           CD := "IEC_Counter_0_DB_1485".Q AND ("Barcode413" > 0) AND "ปุ่มยืนยันหน้า Screen",
                           PV := 5,
                           CV => "Barcode413");
   "M413" := "IEC_Counter_0_DB_440".QU;
   "IEC_Counter_0_DB_1486".CTU(CU := "ยา 414" = 1,
                           R := "Stepper Motor ทำงาน สั่งconveyor เคลื่อที่ไปข้างหน้า" OR "ปุ่มClear",
                           PV := 1);
   "IEC_Counter_0_DB_441".CTUD(CU := ("Expected/Value_All".V = "Expected/Value_All".Expected_414) AND NOT "M414",
                           CD := "IEC_Counter_0_DB_1486".Q AND ("Barcode414" > 0) AND "ปุ่มยืนยันหน้า Screen",
                           PV := 5,
                           CV => "Barcode414");
   "M414" := "IEC_Counter_0_DB_441".QU;
   "IEC_Counter_0_DB_1487".CTU(CU := "ยา 415" = 1,
                           R := "Stepper Motor ทำงาน สั่งconveyor เคลื่อที่ไปข้างหน้า" OR "ปุ่มClear",
                           PV := 1);
   "IEC_Counter_0_DB_442".CTUD(CU := ("Expected/Value_All".V = "Expected/Value_All".Expected_415) AND NOT "M415",
                           CD := "IEC_Counter_0_DB_1487".Q AND ("Barcode415" > 0) AND "ปุ่มยืนยันหน้า Screen",
                           PV := 5,
                           CV => "Barcode415");
   "M415" := "IEC_Counter_0_DB_442".QU;
   "IEC_Counter_0_DB_1488".CTU(CU := "ยา 416" = 1,
                           R := "Stepper Motor ทำงาน สั่งconveyor เคลื่อที่ไปข้างหน้า" OR "ปุ่มClear",
                           PV := 1);
   "IEC_Counter_0_DB_443".CTUD(CU := ("Expected/Value_All".V = "Expected/Value_All".Expected_416) AND NOT "M416",
                           CD := "IEC_Counter_0_DB_1488".Q AND ("Barcode416" > 0) AND "ปุ่มยืนยันหน้า Screen",
                           PV := 5,
                           CV => "Barcode416");
   "M416" := "IEC_Counter_0_DB_443".QU;
   "IEC_Counter_0_DB_1489".CTU(CU := "ยา 417" = 1,
                           R := "Stepper Motor ทำงาน สั่งconveyor เคลื่อที่ไปข้างหน้า" OR "ปุ่มClear",
                           PV := 1);
   "IEC_Counter_0_DB_444".CTUD(CU := ("Expected/Value_All".V = "Expected/Value_All".Expected_417) AND NOT "M417",
                           CD := "IEC_Counter_0_DB_1489".Q AND ("Barcode417" > 0) AND "ปุ่มยืนยันหน้า Screen",
                           PV := 5,
                           CV => "Barcode417");
   "M417" := "IEC_Counter_0_DB_444".QU;
   "IEC_Counter_0_DB_1490".CTU(CU := "ยา 418" = 1,
                           R := "Stepper Motor ทำงาน สั่งconveyor เคลื่อที่ไปข้างหน้า" OR "ปุ่มClear",
                           PV := 1);
   "IEC_Counter_0_DB_445".CTUD(CU := ("Expected/Value_All".V = "Expected/Value_All".Expected_418) AND NOT "M418",
                           CD := "IEC_Counter_0_DB_1490".Q AND ("Barcode418" > 0) AND "ปุ่มยืนยันหน้า Screen",
                           PV := 5,
                           CV => "Barcode418");
   "M418" := "IEC_Counter_0_DB_445".QU;
   "IEC_Counter_0_DB_1491".CTU(CU := "ยา 419" = 1,
                           R := "Stepper Motor ทำงาน สั่งconveyor เคลื่อที่ไปข้างหน้า" OR "ปุ่มClear",
                           PV := 1);
   "IEC_Counter_0_DB_446".CTUD(CU := ("Expected/Value_All".V = "Expected/Value_All".Expected_419) AND NOT "M419",
                           CD := "IEC_Counter_0_DB_1491".Q AND ("Barcode419" > 0) AND "ปุ่มยืนยันหน้า Screen",
                           PV := 5,
                           CV => "Barcode419");
   "M419" := "IEC_Counter_0_DB_446".QU;
   "IEC_Counter_0_DB_1492".CTU(CU := "ยา 420" = 1,
                           R := "Stepper Motor ทำงาน สั่งconveyor เคลื่อที่ไปข้างหน้า" OR "ปุ่มClear",
                           PV := 1);
   "IEC_Counter_0_DB_447".CTUD(CU := ("Expected/Value_All".V = "Expected/Value_All".Expected_420) AND NOT "M420",
                           CD := "IEC_Counter_0_DB_1492".Q AND ("Barcode420" > 0) AND "ปุ่มยืนยันหน้า Screen",
                           PV := 5,
                           CV => "Barcode420");
   "M420" := "IEC_Counter_0_DB_447".QU;
END_REGION

REGION Network 22
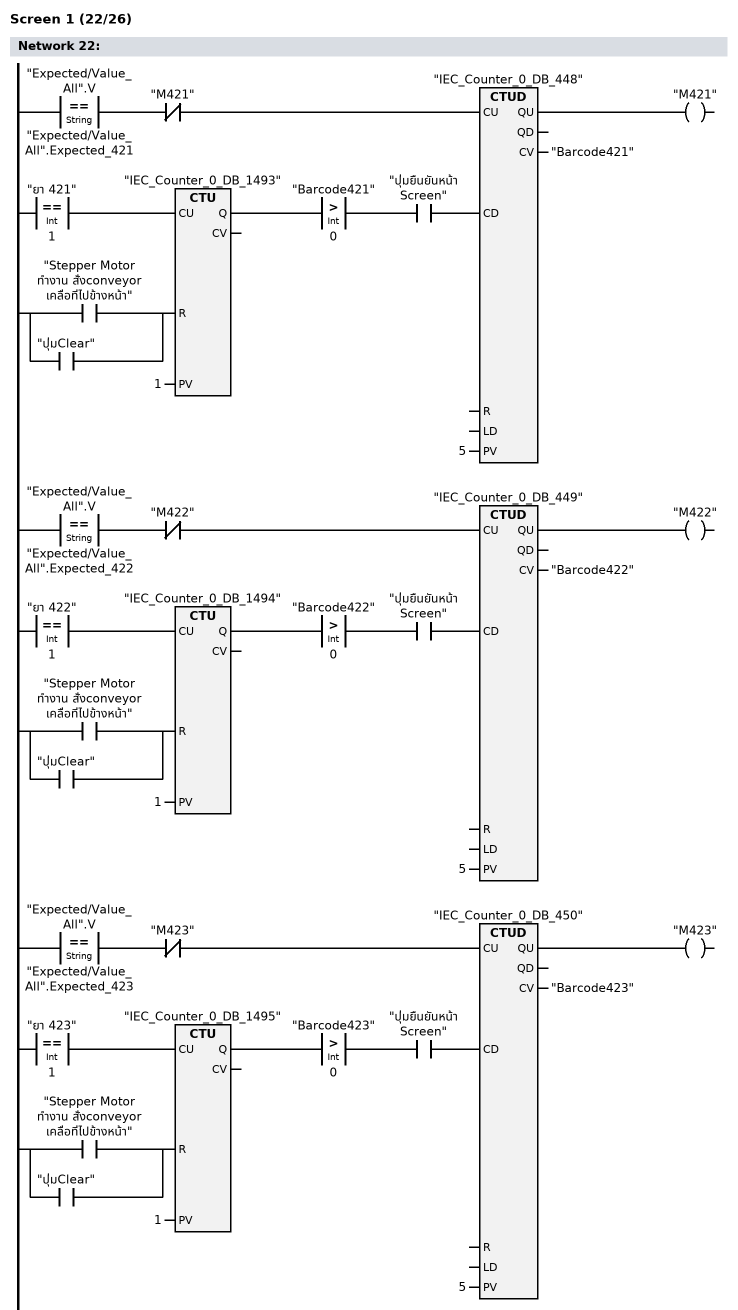
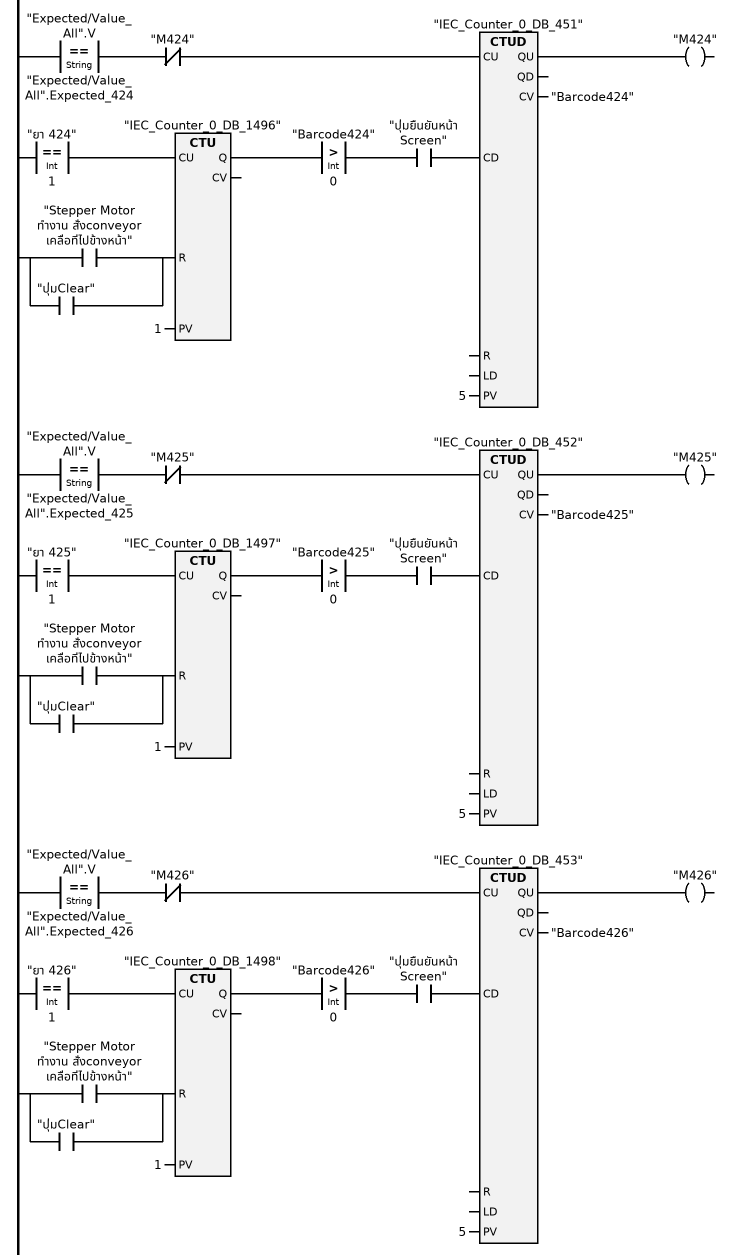
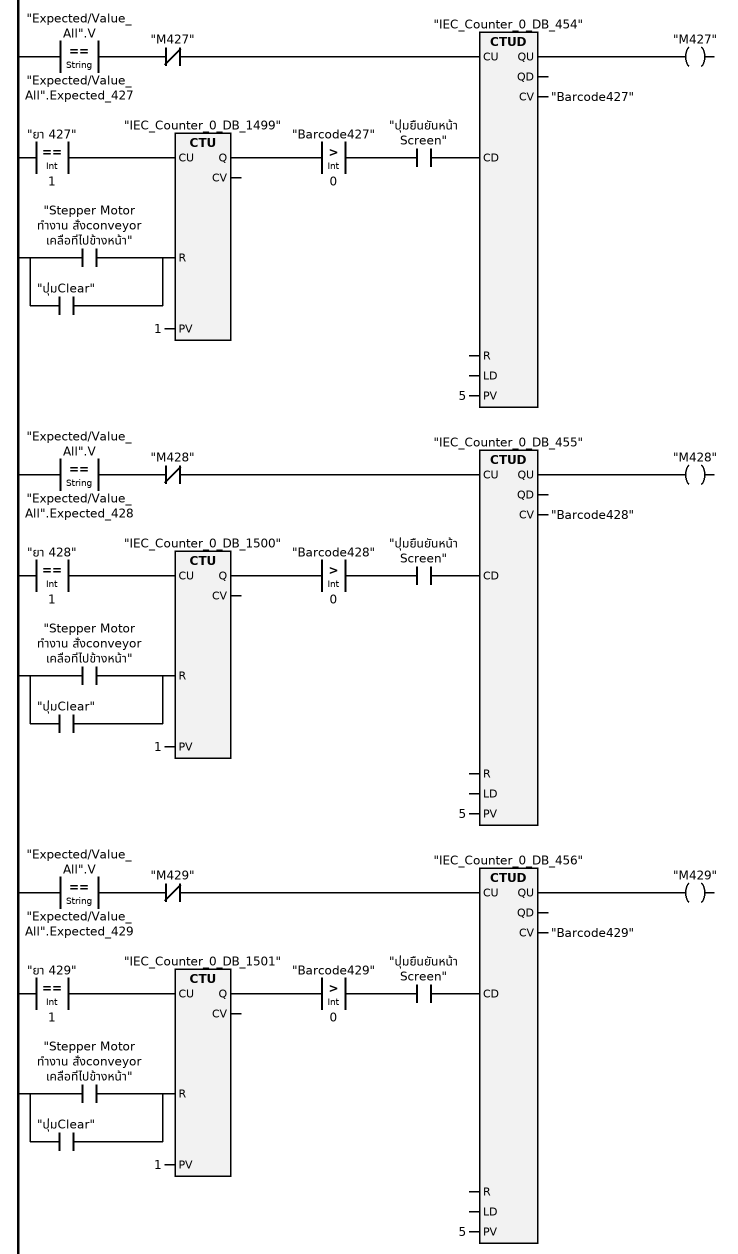
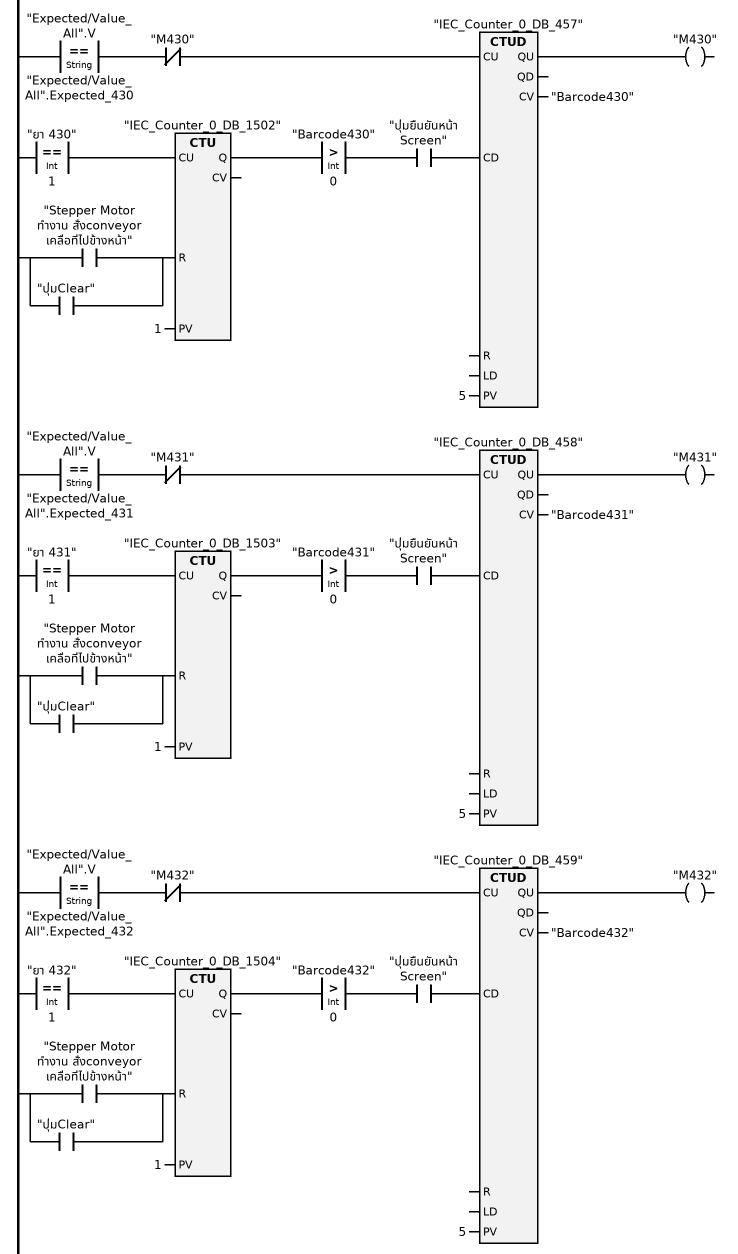
